FUNCTION WRITE_PROTECTED_BYTE
VAR_INPUT
    Ptr : POINTER TO BYTE;
    Value : BYTE;
END_VAR

Ptr^ := Value;

END_FUNCTION

(* stored: Version 1.1.0.1
   POU WRITE_PROTECTED_BYTE: Id {0bd58fcc-2342-4cd5-b054-08bdfb22baa1}, SpecialFunc None *)
